TYPE TcoAbbRW_Inputs_v_8_2_x :
STRUCT
	Inputs AT %I* : ARRAY[0..63] OF BYTE;
END_STRUCT
END_TYPE

(* stored: Version 1.1.0.1, ProductVersion 3.1.4024.12
   DUT TcoAbbRW_Inputs_v_8_2_x: Id {f21766ef-57dd-4f2f-9bf7-65952f4d5e78} *)
